// Mock of FB_DerotatorControl for the telescope state machine tests (MONETcommon#36, BROTLib plan 2026-10-21-telescope-state-machine-unification D1).
FUNCTION_BLOCK FB_DerotatorMock EXTENDS HalfBROT.FB_DerotatorControl
VAR_INPUT
	nMockMoveScans	: UINT := 60;	// scans a move takes (the telescope sees Busy meanwhile)
	bMockLatchTarget	: BOOL;	// #252: a move ends at the target of its start (like MC_MoveAbsolute), not at the current one
	fMockFollowingError	: LREAL;	// #267: deg the encoder lags the NC set position (ActualPosition = SetPosition - this); 0 = none
	nMockStopScans	: UINT := 3;	// scans an MC_Stop takes until Done
	nMockHomeScans	: UINT := 3;	// scans a homing takes
	nMockDisableScans	: UINT := 1;	// scans MC_ExtSetPointGenDisable takes (BROTLib#101)
END_VAR
VAR_OUTPUT
	nStopEdges		: UINT;			// stop requests the telescope made (rising edges of StopAxis)
	nExtErrors		: UINT;			// stop or move requests that met the external setpoint generator (0x4257)
	nResetEdges		: UINT;			// resets the telescope sent to the axis (Reset())
END_VAR
VAR
	fbCore	: FB_AxisMockCore;
	pBool	: POINTER TO BOOL;
	pLreal	: POINTER TO LREAL;
	bInjected	: BOOL;
	nInjectedId	: UDINT;
END_VAR

// No SUPER^(): the real body (MC_* blocks, AXIS_REF) does not run. The real property setters (MoveAxis -> fbAxis.MoveTo(),
// StopAxis -> fbAxis.Stop(), HomeAxis -> _StartHoming) stay, so the telescope sees the real command interface. The model
// is driven by the levels the telescope writes and writes what the telescope reads: the base outputs and, through pointers
// (FB_Axis outputs are not writable from outside), the nested fbAxis outputs.
fbCore(bEnable := bEnable, bHome := bHomeAxis, bMove := bMoveAxis, bStop := bStopAxis, fTarget := fPosition, fHomePosition := fCalibPosition,
	bTracking := bTracking, bLatchTarget := bMockLatchTarget, nMoveScans := nMockMoveScans, nStopScans := nMockStopScans, nHomeScans := nMockHomeScans,
	nDisableScans := nMockDisableScans);

pBool := ADR(fbAxis.Ready);			pBool^ := fbCore.bReady;
pBool := ADR(fbAxis.Calibrated);	pBool^ := fbCore.bCalibrated;
pBool := ADR(fbAxis.HomeDone);		pBool^ := fbCore.bCalibrated;
pBool := ADR(fbAxis.HomeActive);	pBool^ := fbCore.bHoming;
pBool := ADR(fbAxis.Homing);		pBool^ := fbCore.bHoming;
pBool := ADR(fbAxis.InMotion);		pBool^ := fbCore.bInMotion OR fbCore.bTrackActive OR fbCore.bCoast;
pBool := ADR(fbAxis.isTracking);	pBool^ := fbCore.bTrackActive;
pBool := ADR(fbAxis.StandStill);	pBool^ := fbCore.bStandStill AND NOT fbCore.bTrackActive AND NOT fbCore.bCoast;
pBool := ADR(fbAxis.MoveDone);		pBool^ := fbCore.bMoveDone;
pBool := ADR(fbAxis.Stopping);		pBool^ := fbCore.bStopping;
pBool := ADR(fbAxis.StopDone);		pBool^ := fbCore.bStopDone;
pBool := ADR(fbAxis.Busy);			pBool^ := fbCore.bInMotion OR fbCore.bHoming;
pLreal := ADR(fbAxis.ActualPosition);	pLreal^ := fbCore.fPosition - fMockFollowingError;
pLreal := ADR(fbAxis.SetPosition);		pLreal^ := fbCore.fPosition;	// the model position is the NC set position (#267)

bReady := fbCore.bReady AND fbCore.bStandStill;
bCalibrated := fbCore.bCalibrated;
fActualPosition := fbCore.fPosition - fMockFollowingError;
nStopEdges := fbCore.nStopEdges;
nExtErrors := fbCore.nExtErrors;
IF fbCore.bExtError THEN
	bInjected := TRUE;
	nInjectedId := 16#4257;	// Motion commands are not allowed for external setpoint generated axis
END_IF

// the real control body clears the levels like this: the move on MoveDone, the stop on StopDone, the homing request
// once the axis is calibrated and the homing procedure is over
IF fbCore.bMoveDone THEN
	bMoveAxis := FALSE;
END_IF
IF fbCore.bStopDone THEN
	bStopAxis := FALSE;
END_IF
IF fbCore.bCalibrated AND NOT fbCore.bHoming THEN
	bHomeAxis := FALSE;
END_IF
IF bReset THEN
	nResetEdges := nResetEdges + 1;
	bReset := FALSE;	// ResetDone at once
	bInjected := FALSE;
END_IF
bError := bInjected;
nErrorID := nInjectedId;

// the axis reports an error with this id until the telescope resets it (bError/nErrorID are what the telescope reads)
METHOD InjectError
VAR_INPUT
	nId	: UDINT;
END_VAR
bInjected := TRUE;
nInjectedId := nId;
END_METHOD

END_FUNCTION_BLOCK

(* stored: Version 1.1.0.1, ProductVersion 3.1.4024.15
   POU FB_DerotatorMock: Id {a5fdee77-15ca-44ee-96da-486af34b10eb}, SpecialFunc None
   Method InjectError: Id {e037f147-f991-4501-a412-a421f40452ff} *)
